(* IEC 61131-3 sources: kns-port-domestic/targets/astra/src/POUs/Log/F_ZeroPad, 2 files *)

(* ---- F_ZeroPad.decl.st ---- *)
// Назначение: десятичная запись числа с ведущими нулями до uiDigits знаков (поля даты и времени CSV журнала);
//             число длиннее uiDigits — без обрезки.
// Автор:      kr0nsch
// Версия:     0.1.0
// Документ:   docs/DESIGN.md, раздел 9.2
FUNCTION F_ZeroPad : STRING(GVL_Const.LOG_NUM_LEN)
VAR_INPUT
    udiValue : UDINT;               // число
    uiDigits : UINT;                // знаков не меньше
END_VAR
VAR
    uiI : UINT;                     // номер добавляемого нуля
END_VAR

(* ---- F_ZeroPad.impl.st ---- *)
F_ZeroPad := UDINT_TO_STRING(udiValue);
FOR uiI := INT_TO_UINT(LEN(F_ZeroPad)) + 1 TO MIN(uiDigits, INT_TO_UINT(GVL_Const.LOG_NUM_LEN)) DO
    F_ZeroPad := CONCAT('0', F_ZeroPad);
END_FOR
